// TIA Portal V21 export
Screen "Alarms"  1024x768, Number=15, Template=Tpl
  ScreenLayer 
